SUBAPPLICATION FU_Messwerte (* Lesen per Modbus (CLIENT_0_8 pollt selbst alle 500 ms, CNF nach jeder Abfrage), skalieren, auf den lokalen OPC-UA-Server publizieren. *)
  (* Standard: 61499-2; Description: Copyright (c) 2026 Franz Höpfinger This program and the accompanying materials are made available under the terms of the Eclipse Public License 2.0 which is available at https://www.eclipse.org/legal/epl-2.0/ SPDX-License-Identifier: EPL-2.0 *)
  (* Version 1.1, 2026-11-02, Franz Höpfinger, Franz Höpfinger, Skalierung in SubApp FU_Skalierung ausgelagert *)
  (* Version 1.0, 2026-11-02, Franz Höpfinger, Franz Höpfinger, aus FU_Demo_H300 herausgeloest *)
  PACKAGE FBs::FU_Demo;
  IMPORT FBs::FU_Demo::FU_Demo_Konstanten::FU_MODBUS_LESEN;
  IMPORT FBs::FU_Demo::FU_Demo_Konstanten::FU_MESSWERTE_WEB_WRITE;
  FBS
    Lesen : iec61499::net::CLIENT_0_8(QI := TRUE, ID := FU_MODBUS_LESEN); (* 9000H..9004H, 9006H, 9332H, 9333H. Pollt selbst (pollFrequency 500 ms im ID-String) und loest nach jeder erfolgreichen Abfrage CNF aus - kein REQ, kein E_CYCLE noetig. *)
    Publish_Messwerte : iec61499::net::PUBLISH_8(QI := TRUE, ID := FU_MESSWERTE_WEB_WRITE);
  END_FBS
  SUBAPPS
    Skalierung : FBs::FU_Demo::FU_Skalierung;
  END_SUBAPPS
  EVENT_CONNECTIONS
    Lesen.CNF TO Skalierung.REQ;
    Skalierung.CNF TO Publish_Messwerte.REQ;
  END_CONNECTIONS
  DATA_CONNECTIONS
    Lesen.RD_1 TO Skalierung.RD_1;
    Lesen.RD_2 TO Skalierung.RD_2;
    Lesen.RD_3 TO Skalierung.RD_3;
    Lesen.RD_4 TO Skalierung.RD_4;
    Lesen.RD_5 TO Skalierung.RD_5;
    Lesen.RD_6 TO Skalierung.RD_6;
    Lesen.RD_7 TO Skalierung.RD_7;
    Lesen.RD_8 TO Skalierung.RD_8;
    Skalierung.SD_1 TO Publish_Messwerte.SD_1;
    Skalierung.SD_2 TO Publish_Messwerte.SD_2;
    Skalierung.SD_3 TO Publish_Messwerte.SD_3;
    Skalierung.SD_4 TO Publish_Messwerte.SD_4;
    Skalierung.SD_5 TO Publish_Messwerte.SD_5;
    Skalierung.SD_6 TO Publish_Messwerte.SD_6;
    Skalierung.SD_7 TO Publish_Messwerte.SD_7;
    Skalierung.SD_8 TO Publish_Messwerte.SD_8;
  END_CONNECTIONS
END_SUBAPPLICATION
